PROGRAM main
  VAR
    SCADA_HVAC_RAIL_CMD AT %QX0.0 : BOOL;
    SCADA_FIRE_RAIL_CMD AT %QX0.1 : BOOL;
    SCADA_DOOR_RAIL_CMD AT %QX0.2 : BOOL;
    PUB_HVAC_RAIL_STATUS AT %QX0.3 : BOOL;
    PUB_FIRE_RAIL_STATUS AT %QX0.4 : BOOL;
    PUB_DOOR_RAIL_STATUS AT %QX0.5 : BOOL;
    PUB_HEARTBEAT AT %QW0 : UINT;
    PUB_RECONNECT_COUNT AT %QW1 : UINT;
    HVAC_RAIL_CMD AT %QX100.0 : BOOL;
    FIRE_RAIL_CMD AT %QX100.1 : BOOL;
    DOOR_RAIL_CMD AT %QX100.2 : BOOL;
    HVAC_RAIL_STATUS AT %IX100.0 : BOOL;
    FIRE_RAIL_STATUS AT %IX100.1 : BOOL;
    DOOR_RAIL_STATUS AT %IX100.2 : BOOL;
    HEARTBEAT AT %IW100 : UINT;
    RECONNECT_COUNT AT %IW101 : UINT;
  END_VAR

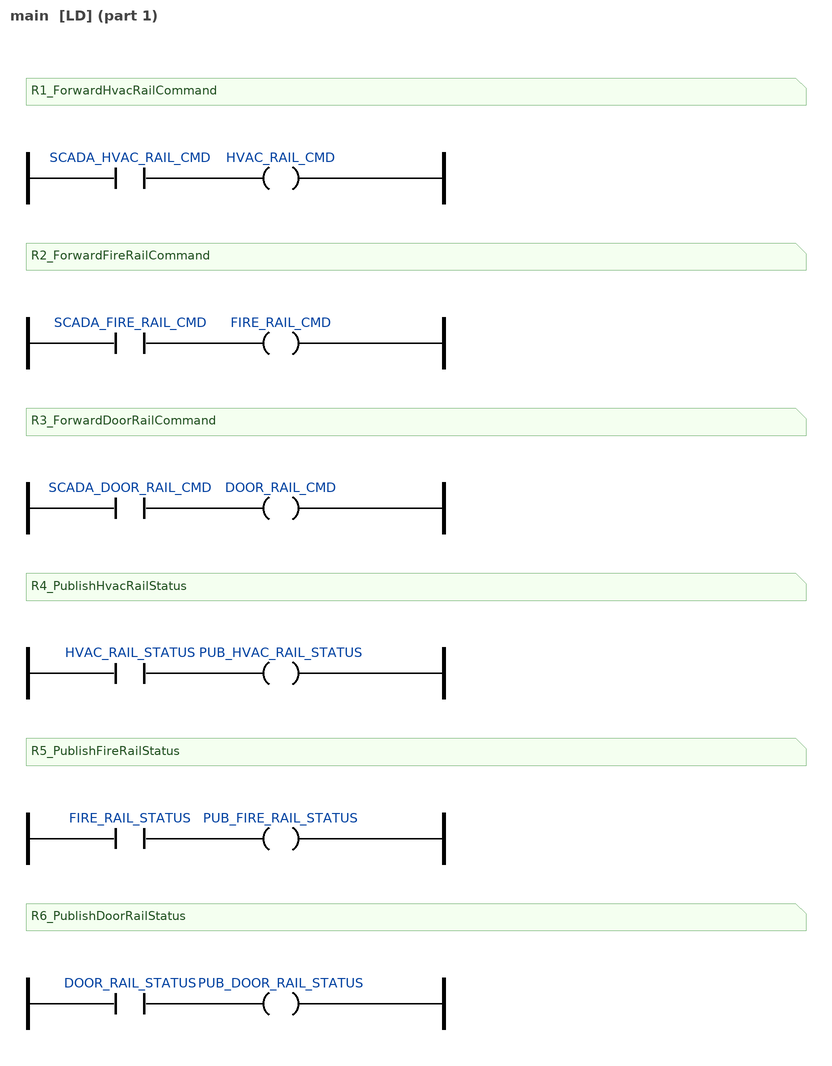
(* LD diagram, written out as Structured Text *)
(* R1_ForwardHvacRailCommand *)
HVAC_RAIL_CMD := SCADA_HVAC_RAIL_CMD;
(* R2_ForwardFireRailCommand *)
FIRE_RAIL_CMD := SCADA_FIRE_RAIL_CMD;
(* R3_ForwardDoorRailCommand *)
DOOR_RAIL_CMD := SCADA_DOOR_RAIL_CMD;
(* R4_PublishHvacRailStatus *)
PUB_HVAC_RAIL_STATUS := HVAC_RAIL_STATUS;
(* R5_PublishFireRailStatus *)
PUB_FIRE_RAIL_STATUS := FIRE_RAIL_STATUS;
(* R6_PublishDoorRailStatus *)
PUB_DOOR_RAIL_STATUS := DOOR_RAIL_STATUS;
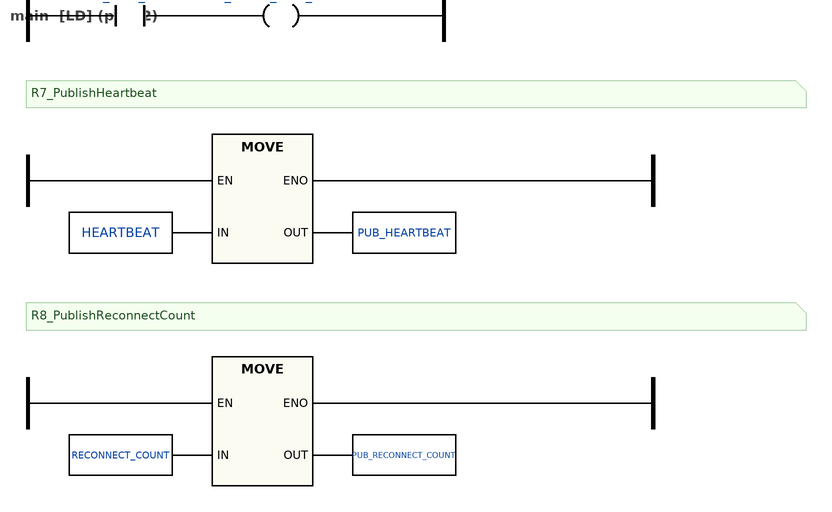
(* R7_PublishHeartbeat *)
PUB_HEARTBEAT := HEARTBEAT;
(* R8_PublishReconnectCount *)
PUB_RECONNECT_COUNT := RECONNECT_COUNT;
END_PROGRAM
